SUBAPPLICATION GreenRedBackground2SC (* Hintergrundfarbe (TRUE -> Grün, FALSE -> Rot) für 2 Objekte (Kompakt) *)
  (* Standard: 61499-2 *)
  (* Version 1.0, 2026-07-21, franz, Meisterschulen am Ostbahnhof *)
  PACKAGE MyLib::sys;
  IMPORT isobus::UT::Q::types::s2ObjectIDs;
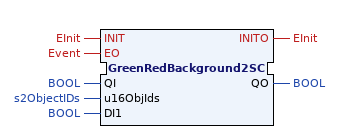
  EVENT_INPUT
    INIT : EInit; (* Initialization Request *)
    EO;
  END_EVENT
  EVENT_OUTPUT
    INITO : EInit; (* Initialization Confirm *)
  END_EVENT
  VAR_INPUT
    QI : BOOL := TRUE; (* Quality Input - TRUE to enable service *)
    u16ObjIds : isobus::UT::Q::types::s2ObjectIDs;
    DI1 : BOOL; (* Selector *)
  END_VAR
  VAR_OUTPUT
    QO : BOOL; (* Quality Output - TRUE if service executed successfully *)
  END_VAR
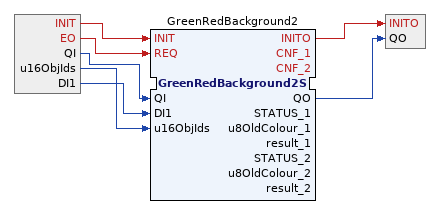
  SUBAPPS
    GreenRedBackground2 : MyLib::sys::GreenRedBackground2S;
  END_SUBAPPS
  EVENT_CONNECTIONS
    EO TO GreenRedBackground2.REQ;
    INIT TO GreenRedBackground2.INIT;
    GreenRedBackground2.INITO TO INITO;
  END_CONNECTIONS
  DATA_CONNECTIONS
    u16ObjIds TO GreenRedBackground2.u16ObjIds;
    DI1 TO GreenRedBackground2.DI1;
    QI TO GreenRedBackground2.QI;
    GreenRedBackground2.QO TO QO;
  END_CONNECTIONS
END_SUBAPPLICATION
